Fanuc KAREL source: ka00165.KL

-- PROVISIONAL review KL for V1013-1; original PC SHA256 96e172bf694b5d1bf729d803a6386270fc552716b3297b644fd9cc0491677ab8
-- Incomplete behavior may be omitted. Consult companion uncertainty JSON. Do not deploy.
PROGRAM KA00165
%NOLOCKGROUP
-- UNRESOLVED_DECL SRC type=002012
-- UNRESOLVED_DECL DST type=002012
BEGIN
  -- UNRESOLVED_PC offsets 5-19; opcodes 22,22,1E
  -- UNRESOLVED_PC offsets 24-28; opcodes 7F
END KA00165
